(* PLC project Pump station (ladder), Digital twin lab Pump station 1 *)
(* stored: creationDateTime 2026-10-06T00:00:00, modificationDateTime 2026-10-06T00:00:00 *)

(* Lead/lag pump station control in ladder logic. Same behavior, variables and addresses as pump_station.st. *)
PROGRAM PumpStation
  VAR
    P1_RUNNING AT %IX100.0 : BOOL;  (* P1 running feedback (simulator DI 0) *)
    P2_RUNNING AT %IX100.1 : BOOL;  (* P2 running feedback (simulator DI 1) *)
    P1_FAULT AT %IX100.2 : BOOL;  (* P1 fault / trip (simulator DI 2) *)
    P2_FAULT AT %IX100.3 : BOOL;  (* P2 fault / trip (simulator DI 3) *)
    PT101_DISCH AT %IW100 : UINT;  (* Discharge pressure PT-101, psi x10 *)
    PT100_SUCT AT %IW101 : UINT;  (* Suction pressure PT-100, psi x10 *)
    DEMAND AT %IW102 : UINT;  (* Pipeline demand, % x10 *)
    SIM_HEARTBEAT AT %IW103 : UINT;  (* Simulator heartbeat, +1 every simulator step *)
    P1_RUN_CMD AT %QX100.0 : BOOL;  (* P1 run command (simulator coil 0) *)
    P2_RUN_CMD AT %QX100.1 : BOOL;  (* P2 run command (simulator coil 1) *)
    HMI_DISCH_PRESS AT %QW0 : UINT;  (* HR 0: discharge pressure, psi x10 *)
    HMI_SUCT_PRESS AT %QW1 : UINT;  (* HR 1: suction pressure, psi x10 *)
    HMI_DEMAND AT %QW2 : UINT;  (* HR 2: demand, % x10 *)
    HMI_STATUS AT %QW3 : UINT;  (* HR 3: status bits (design 5.2) *)
    HMI_ALARMS AT %QW4 : UINT;  (* HR 4: alarm bits (design 5.2) *)
    HMI_LEAD_PUMP AT %QW5 : UINT;  (* HR 5: active lead pump, 1 or 2 *)
    HMI_MODE_ACTIVE AT %QW6 : UINT;  (* HR 6: active mode, 0 Off 1 Auto 2 Manual *)
    PLC_HEARTBEAT AT %QW7 : UINT;  (* HR 7: +1 every PLC scan *)
    SP_PRESSURE AT %MW0 : UINT;  (* HR 1024: lag start pressure, psi x10 *)
    SP_LAG_STOP AT %MW1 : UINT;  (* HR 1025: lag stop pressure, psi x10 *)
    SP_LOW_ALARM AT %MW2 : UINT;  (* HR 1026: low pressure alarm, psi x10 *)
    SP_HIGH_ALARM AT %MW3 : UINT;  (* HR 1027: high pressure alarm, psi x10 *)
    LAG_START_DELAY AT %MW4 : UINT;  (* HR 1028: lag start delay, s *)
    LAG_STOP_DELAY AT %MW5 : UINT;  (* HR 1029: lag stop delay, s *)
    CMD_MODE AT %MW6 : UINT;  (* HR 1030: mode command, 0 Off 1 Auto 2 Manual *)
    CMD_LEAD_SELECT AT %MW7 : UINT;  (* HR 1031: lead pump select, 1 = P1, 2 = P2 *)
    CMD_MANUAL_P1 AT %MW8 : UINT;  (* HR 1032: Manual mode P1, 1 run 0 stop *)
    CMD_MANUAL_P2 AT %MW9 : UINT;  (* HR 1033: Manual mode P2, 1 run 0 stop *)
    CMD_ALARM_RESET AT %MW10 : UINT;  (* HR 1034: alarm reset, HMI writes 1, PLC clears it *)
  END_VAR
  VAR
    LoadDefaults : BOOL;  (* SP_PRESSURE is 0: settings were never written, load defaults *)
    MinLagStop : UINT;  (* SP_PRESSURE + 10 psi, the lowest allowed lag stop pressure *)
    ModeAuto : BOOL;  (* CMD_MODE = 1 *)
    ModeManual : BOOL;  (* CMD_MODE = 2 *)
    SelP2 : BOOL;  (* CMD_LEAD_SELECT = 2 (operator wants P2 as lead) *)
    ManP1 : BOOL;  (* CMD_MANUAL_P1 = 1 *)
    ManP2 : BOOL;  (* CMD_MANUAL_P2 = 1 *)
    ResetReq : BOOL;  (* Operator pressed Reset (CMD_ALARM_RESET <> 0) *)
    PressBelowSP : BOOL;  (* Discharge pressure below the lag start pressure *)
    PressAboveLagStop : BOOL;  (* Discharge pressure above the lag stop pressure *)
    PressBelowLowAlm : BOOL;  (* Discharge pressure below the low alarm limit *)
    PressAboveHighAlm : BOOL;  (* Discharge pressure above the high alarm limit *)
    P1StartTmr : TON;  (* P1 commanded but not running *)
    P2StartTmr : TON;  (* P2 commanded but not running *)
    P1StartFail : BOOL;  (* P1 failed to start within 5 s *)
    P2StartFail : BOOL;  (* P2 failed to start within 5 s *)
    P1Failed : BOOL;  (* P1 locked out (fault or failed to start) until Reset *)
    P2Failed : BOOL;  (* P2 locked out (fault or failed to start) until Reset *)
    EnterAuto : BOOL;  (* First scan in Auto *)
    LeadIsP2 : BOOL;  (* Active lead pump: FALSE = P1, TRUE = P2 (ActiveLead in the ST program) *)
    LagPumpCmd : BOOL;  (* The pump that is now lag is commanded to run *)
    FailToP2 : BOOL;  (* Lead P1 has failed and P2 is healthy: make P2 lead *)
    FailToP1 : BOOL;  (* Lead P2 has failed and P1 is healthy: make P1 lead *)
    LeadChange : BOOL;  (* Apply the operator's new lead selection this scan *)
    LagRun : BOOL;  (* Auto logic wants the lag pump running *)
    Handover : BOOL;  (* Lead change in progress: old lead keeps running until the new one runs *)
    LeadAvail : BOOL;  (* Lead pump is not locked out *)
    LagAvail : BOOL;  (* Lag pump is not locked out *)
    LeadRunning : BOOL;  (* Lead pump reports running *)
    LagStartPT : TIME;  (* Lag start delay as TIME *)
    LagStopPT : TIME;  (* Lag stop delay as TIME *)
    LagStartTmr : TON;  (* Pressure low long enough to start the lag pump *)
    LagStopTmr : TON;  (* Pressure high long enough to stop the lag pump *)
    LagStartDone : BOOL;  (* LagStartTmr.Q *)
    LagStopDone : BOOL;  (* LagStopTmr.Q *)
    LowArmTmr : TON;  (* Start-up bypass for the low pressure alarm *)
    LowPressTmr : TON;  (* Low pressure alarm delay *)
    HighPressTmr : TON;  (* High pressure alarm delay *)
    CommLossTmr : TON;  (* Simulator heartbeat frozen *)
    LowArmed : BOOL;  (* Low pressure alarm armed (15 s out of Off) *)
    LowPressOn : BOOL;  (* Pressure low for 5 s *)
    HighPressOn : BOOL;  (* Pressure high for 5 s *)
    SimHbFrozen : BOOL;  (* Simulator heartbeat unchanged since the last scan *)
    LastSimHb : UINT;  (* Simulator heartbeat seen last scan *)
    CommLost : BOOL;  (* Simulator heartbeat frozen for 3 s *)
    CommOk : BOOL;  (* Simulator link healthy *)
    AlmLow : BOOL;  (* Low discharge pressure alarm (latched) *)
    AlmHigh : BOOL;  (* High discharge pressure alarm (latched) *)
    AlmComm : BOOL;  (* Simulator comm loss alarm (latched) *)
    AlmUnack : BOOL;  (* A new alarm has not been acknowledged *)
    AnyAlarm : BOOL;  (* Any alarm or pump lockout active *)
    LagRunning : BOOL;  (* Lag pump reports running *)
    StatusWord : UINT;  (* HMI_STATUS being built *)
    AlarmWord : UINT;  (* HMI_ALARMS being built *)
    HbWrap : BOOL;  (* PLC_HEARTBEAT is at 65535 and wraps to 0 *)
  END_VAR
  VAR  (* added by the conversion: wires and edge detectors of the diagram *)
    R_TRIG1 : R_TRIG;
    R_TRIG2 : R_TRIG;
  END_VAR

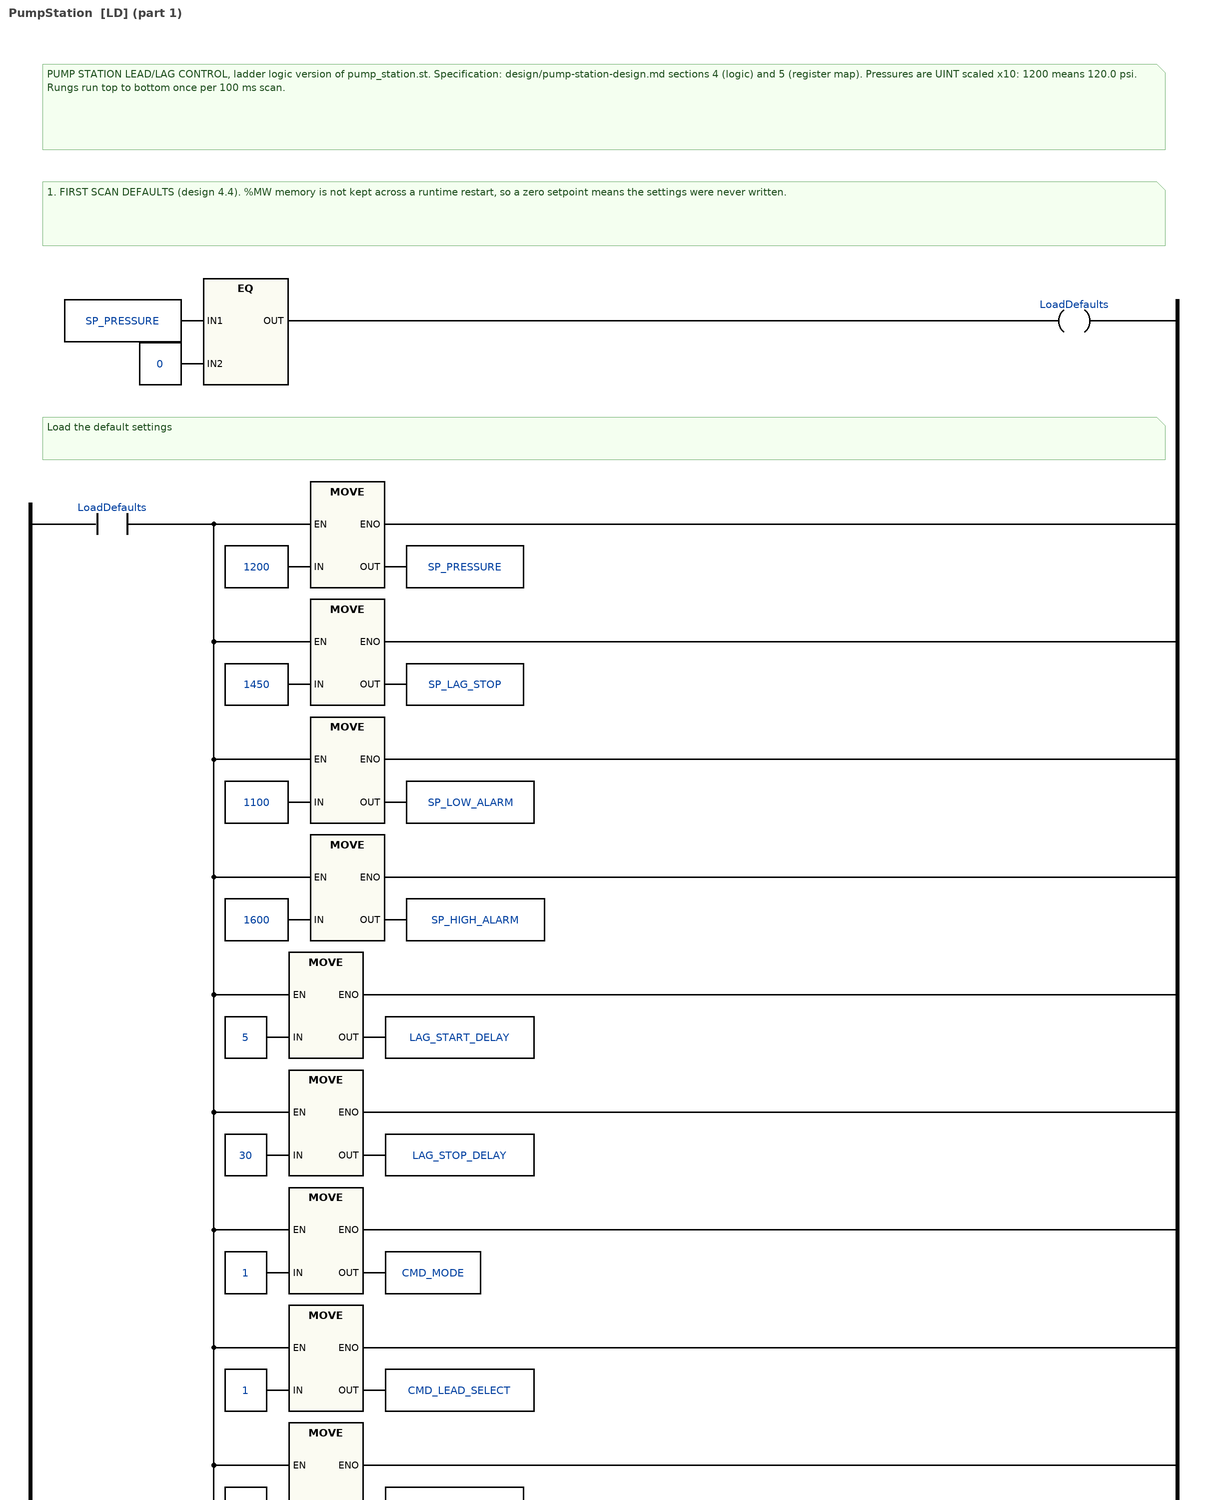
(* LD diagram, written out as Structured Text *)
(* PUMP STATION LEAD/LAG CONTROL, ladder logic version of pump_station.st. Specification: design/pump-station-design.md sections 4 (logic) and 5 (register map). Pressures are UINT scaled x10: 1200 means 120.0 psi. Rungs run top to bottom once per 100 ms scan. *)
(* 1. FIRST SCAN DEFAULTS (design 4.4). %MW memory is not kept across a runtime restart, so a zero setpoint means the settings were never written. *)
LoadDefaults := SP_PRESSURE = 0;
(* Load the default settings *)
IF LoadDefaults THEN SP_PRESSURE := 1200; END_IF;
IF LoadDefaults THEN SP_LAG_STOP := 1450; END_IF;
IF LoadDefaults THEN SP_LOW_ALARM := 1100; END_IF;
IF LoadDefaults THEN SP_HIGH_ALARM := 1600; END_IF;
IF LoadDefaults THEN LAG_START_DELAY := 5; END_IF;
IF LoadDefaults THEN LAG_STOP_DELAY := 30; END_IF;
IF LoadDefaults THEN CMD_MODE := 1; END_IF;
IF LoadDefaults THEN CMD_LEAD_SELECT := 1; END_IF;
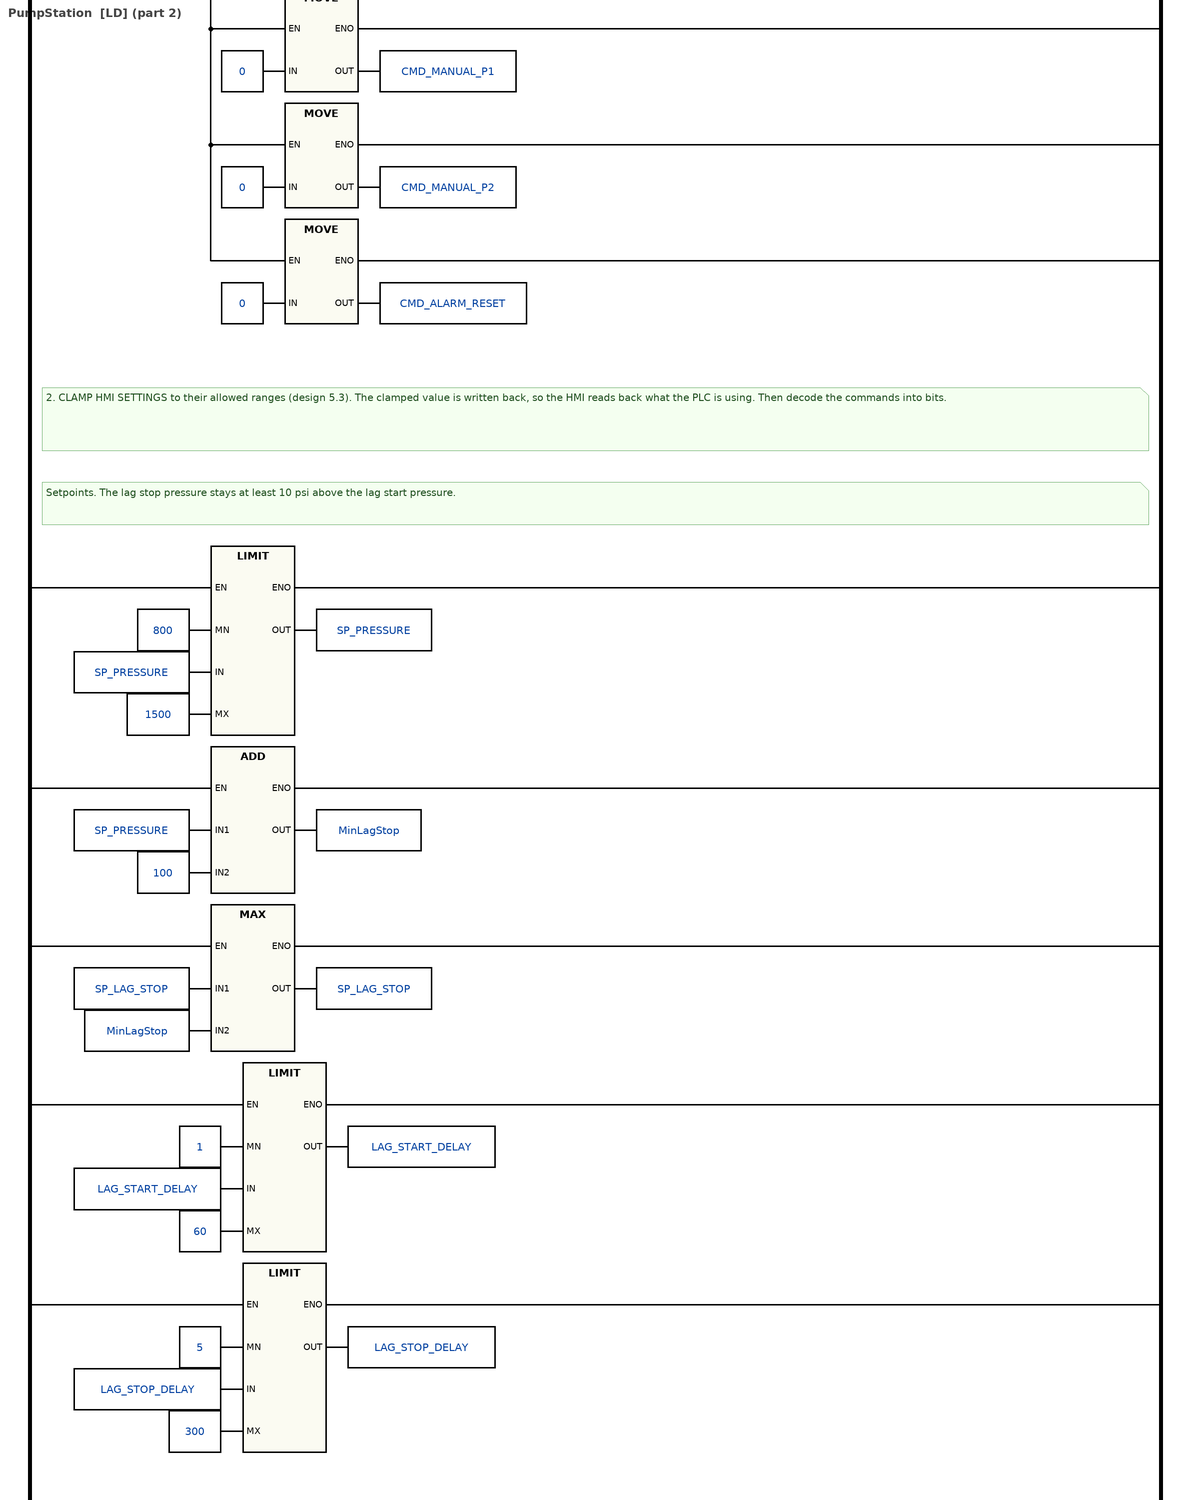
IF LoadDefaults THEN CMD_MANUAL_P1 := 0; END_IF;
IF LoadDefaults THEN CMD_MANUAL_P2 := 0; END_IF;
IF LoadDefaults THEN CMD_ALARM_RESET := 0; END_IF;
(* 2. CLAMP HMI SETTINGS to their allowed ranges (design 5.3). The clamped value is written back, so the HMI reads back what the PLC is using. Then decode the commands into bits. *)
(* Setpoints. The lag stop pressure stays at least 10 psi above the lag start pressure. *)
SP_PRESSURE := LIMIT(800, SP_PRESSURE, 1500);
MinLagStop := SP_PRESSURE + 100;
SP_LAG_STOP := MAX(SP_LAG_STOP, MinLagStop);
LAG_START_DELAY := LIMIT(1, LAG_START_DELAY, 60);
LAG_STOP_DELAY := LIMIT(5, LAG_STOP_DELAY, 300);
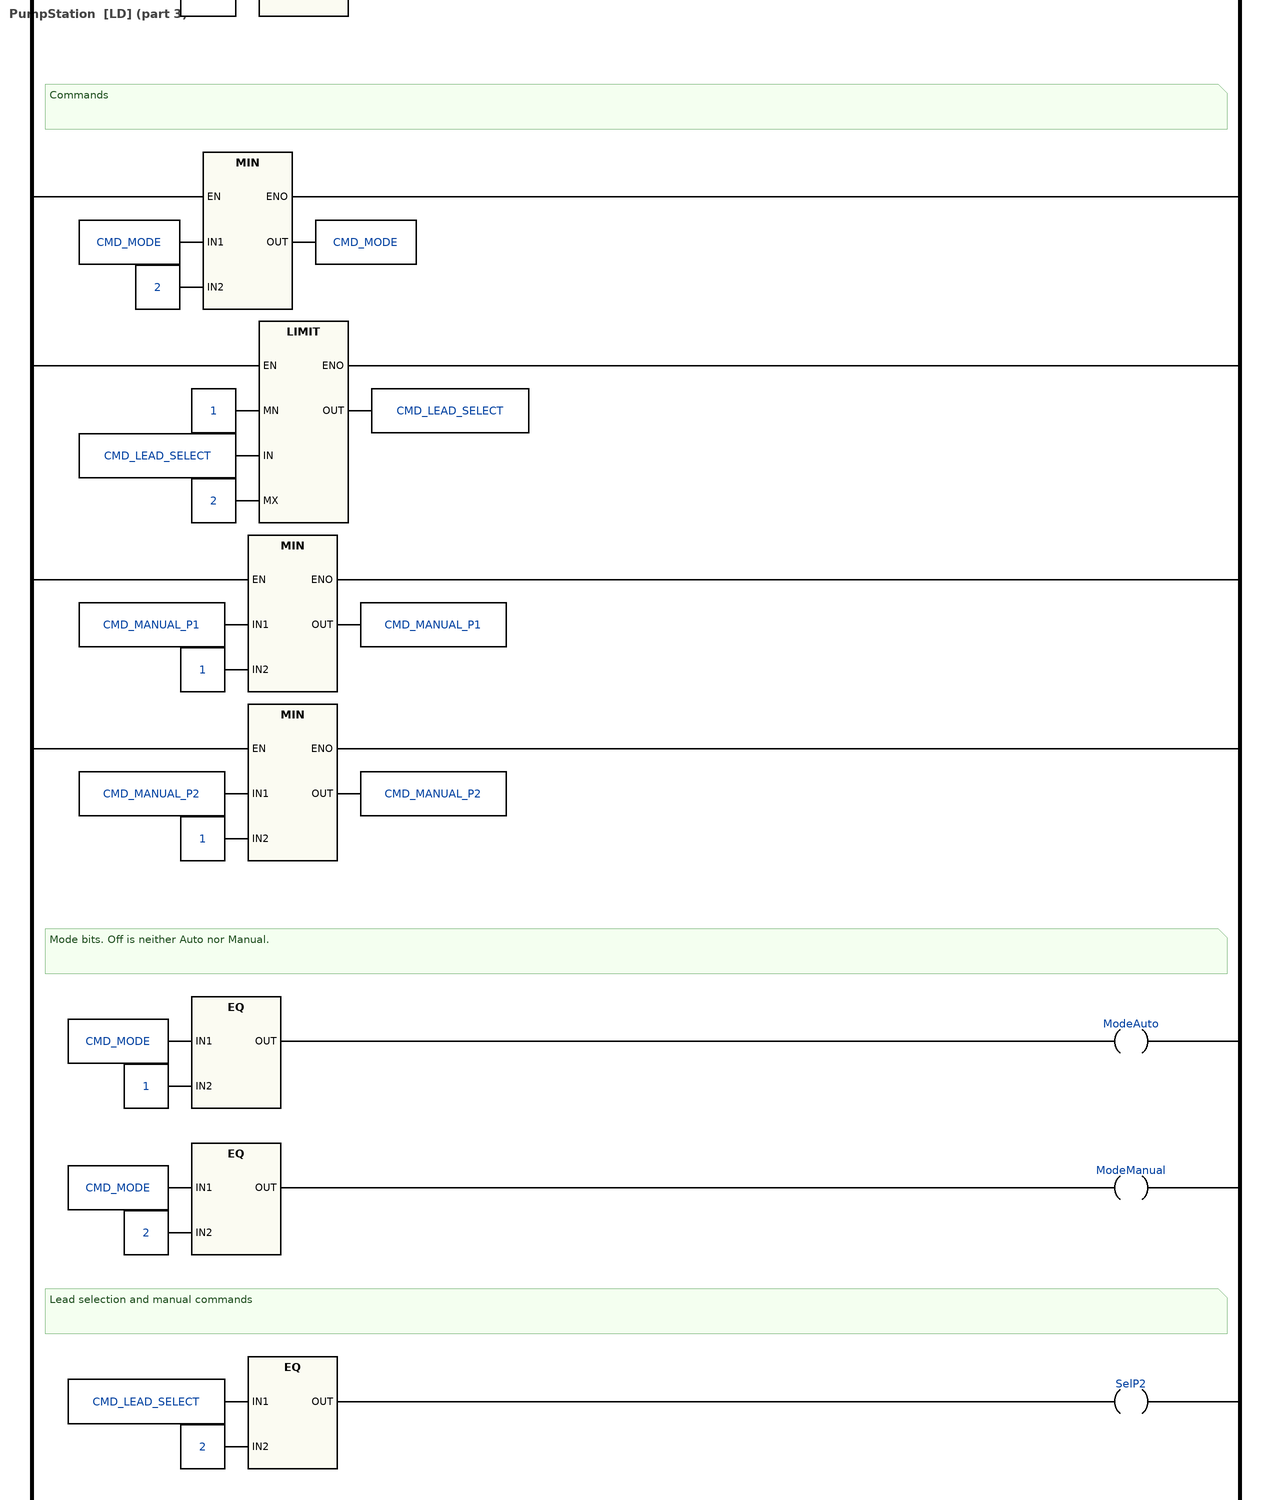
(* Commands *)
CMD_MODE := MIN(CMD_MODE, 2);
CMD_LEAD_SELECT := LIMIT(1, CMD_LEAD_SELECT, 2);
CMD_MANUAL_P1 := MIN(CMD_MANUAL_P1, 1);
CMD_MANUAL_P2 := MIN(CMD_MANUAL_P2, 1);
(* Mode bits. Off is neither Auto nor Manual. *)
ModeAuto := CMD_MODE = 1;
ModeManual := CMD_MODE = 2;
(* Lead selection and manual commands *)
SelP2 := CMD_LEAD_SELECT = 2;
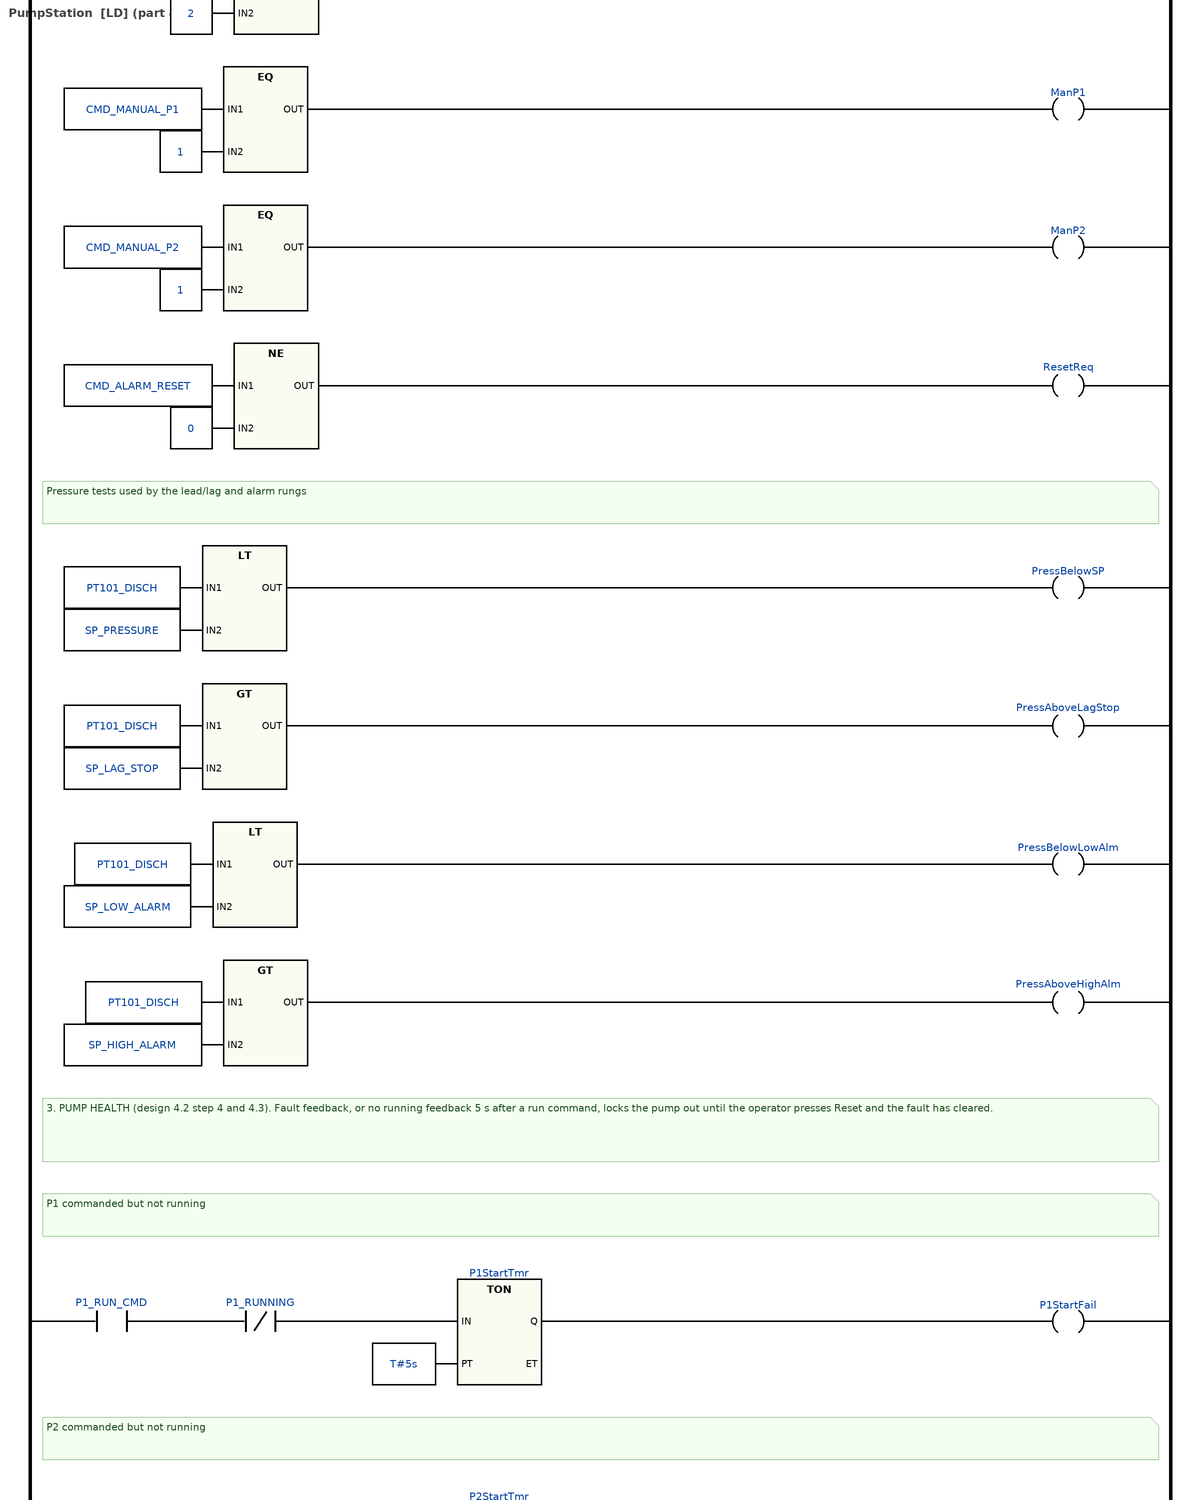
ManP1 := CMD_MANUAL_P1 = 1;
ManP2 := CMD_MANUAL_P2 = 1;
ResetReq := CMD_ALARM_RESET <> 0;
(* Pressure tests used by the lead/lag and alarm rungs *)
PressBelowSP := PT101_DISCH < SP_PRESSURE;
PressAboveLagStop := PT101_DISCH > SP_LAG_STOP;
PressBelowLowAlm := PT101_DISCH < SP_LOW_ALARM;
PressAboveHighAlm := PT101_DISCH > SP_HIGH_ALARM;
(* 3. PUMP HEALTH (design 4.2 step 4 and 4.3). Fault feedback, or no running feedback 5 s after a run command, locks the pump out until the operator presses Reset and the fault has cleared. *)
(* P1 commanded but not running *)
P1StartTmr(IN := P1_RUN_CMD AND NOT P1_RUNNING, PT := T#5s);
P1StartFail := P1StartTmr.Q;
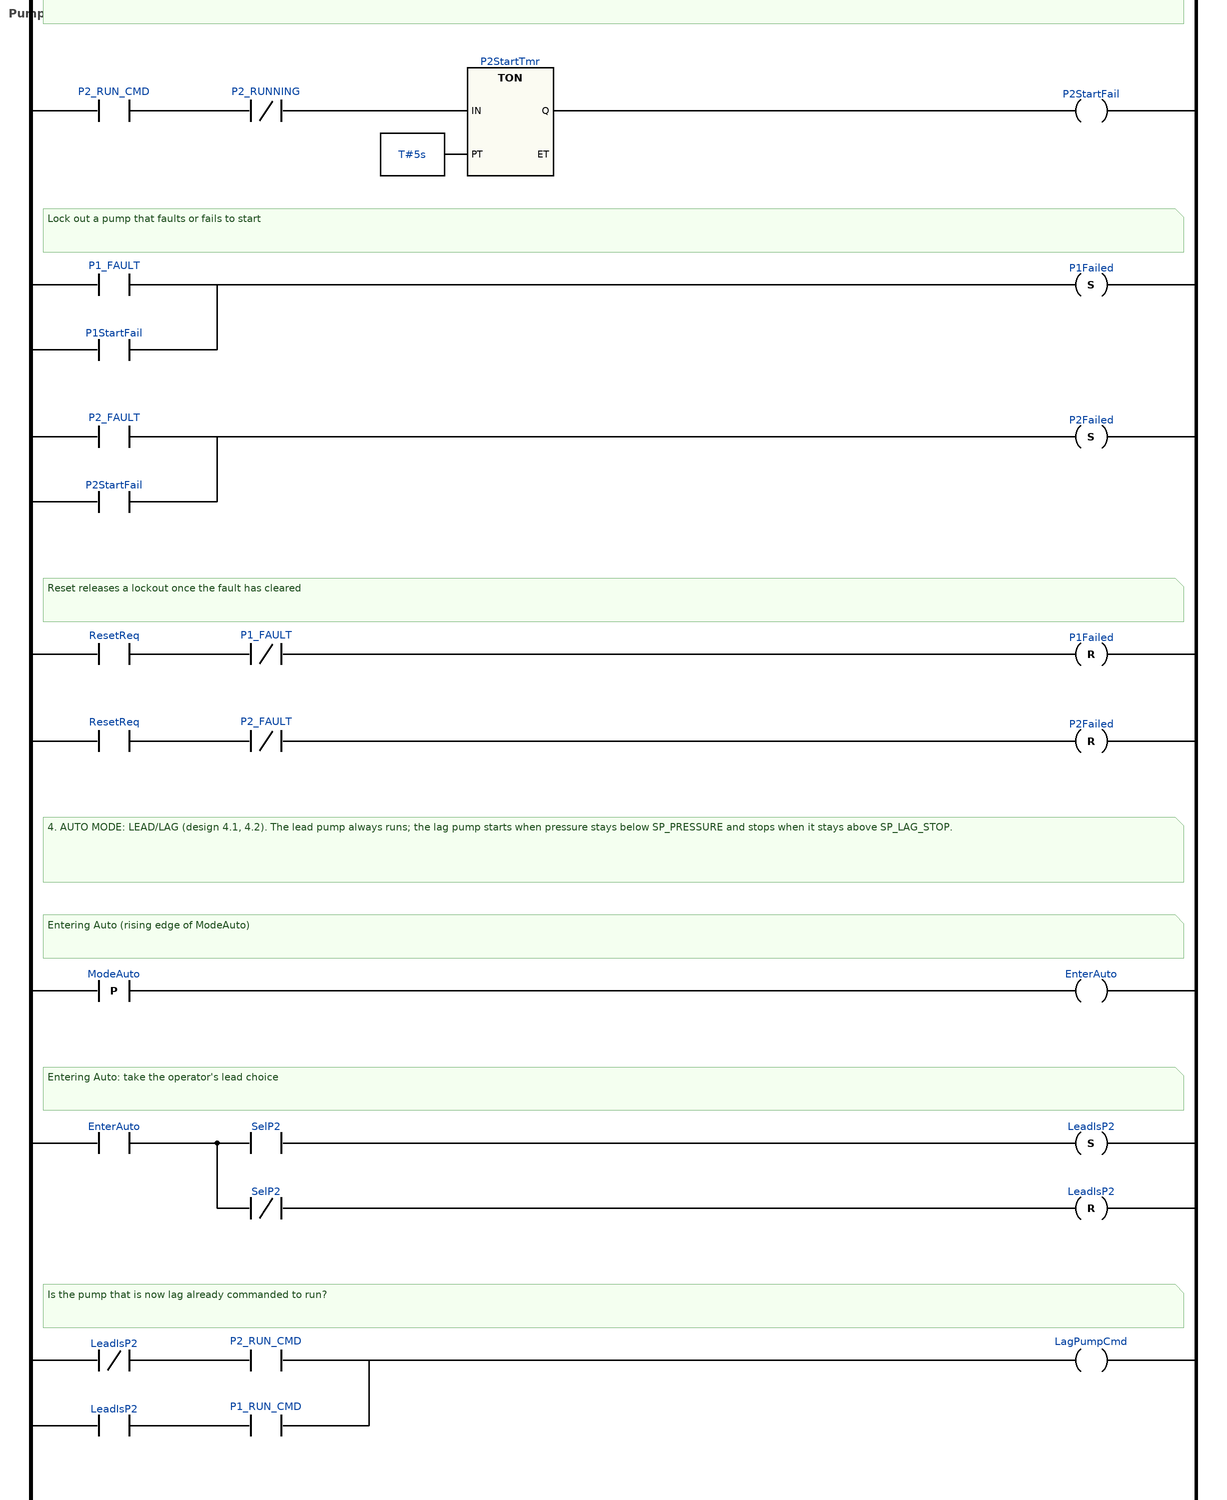
(* P2 commanded but not running *)
P2StartTmr(IN := P2_RUN_CMD AND NOT P2_RUNNING, PT := T#5s);
P2StartFail := P2StartTmr.Q;
(* Lock out a pump that faults or fails to start *)
IF P1_FAULT OR P1StartFail THEN P1Failed := TRUE; END_IF;
IF P2_FAULT OR P2StartFail THEN P2Failed := TRUE; END_IF;
(* Reset releases a lockout once the fault has cleared *)
IF ResetReq AND NOT P1_FAULT THEN P1Failed := FALSE; END_IF;
IF ResetReq AND NOT P2_FAULT THEN P2Failed := FALSE; END_IF;
(* 4. AUTO MODE: LEAD/LAG (design 4.1, 4.2). The lead pump always runs; the lag pump starts when pressure stays below SP_PRESSURE and stops when it stays above SP_LAG_STOP. *)
(* Entering Auto (rising edge of ModeAuto) *)
R_TRIG1(CLK := ModeAuto);
EnterAuto := R_TRIG1.Q;
(* Entering Auto: take the operator's lead choice *)
IF EnterAuto AND SelP2 THEN LeadIsP2 := TRUE; END_IF;
IF EnterAuto AND NOT SelP2 THEN LeadIsP2 := FALSE; END_IF;
(* Is the pump that is now lag already commanded to run? *)
LagPumpCmd := NOT LeadIsP2 AND P2_RUN_CMD OR LeadIsP2 AND P1_RUN_CMD;
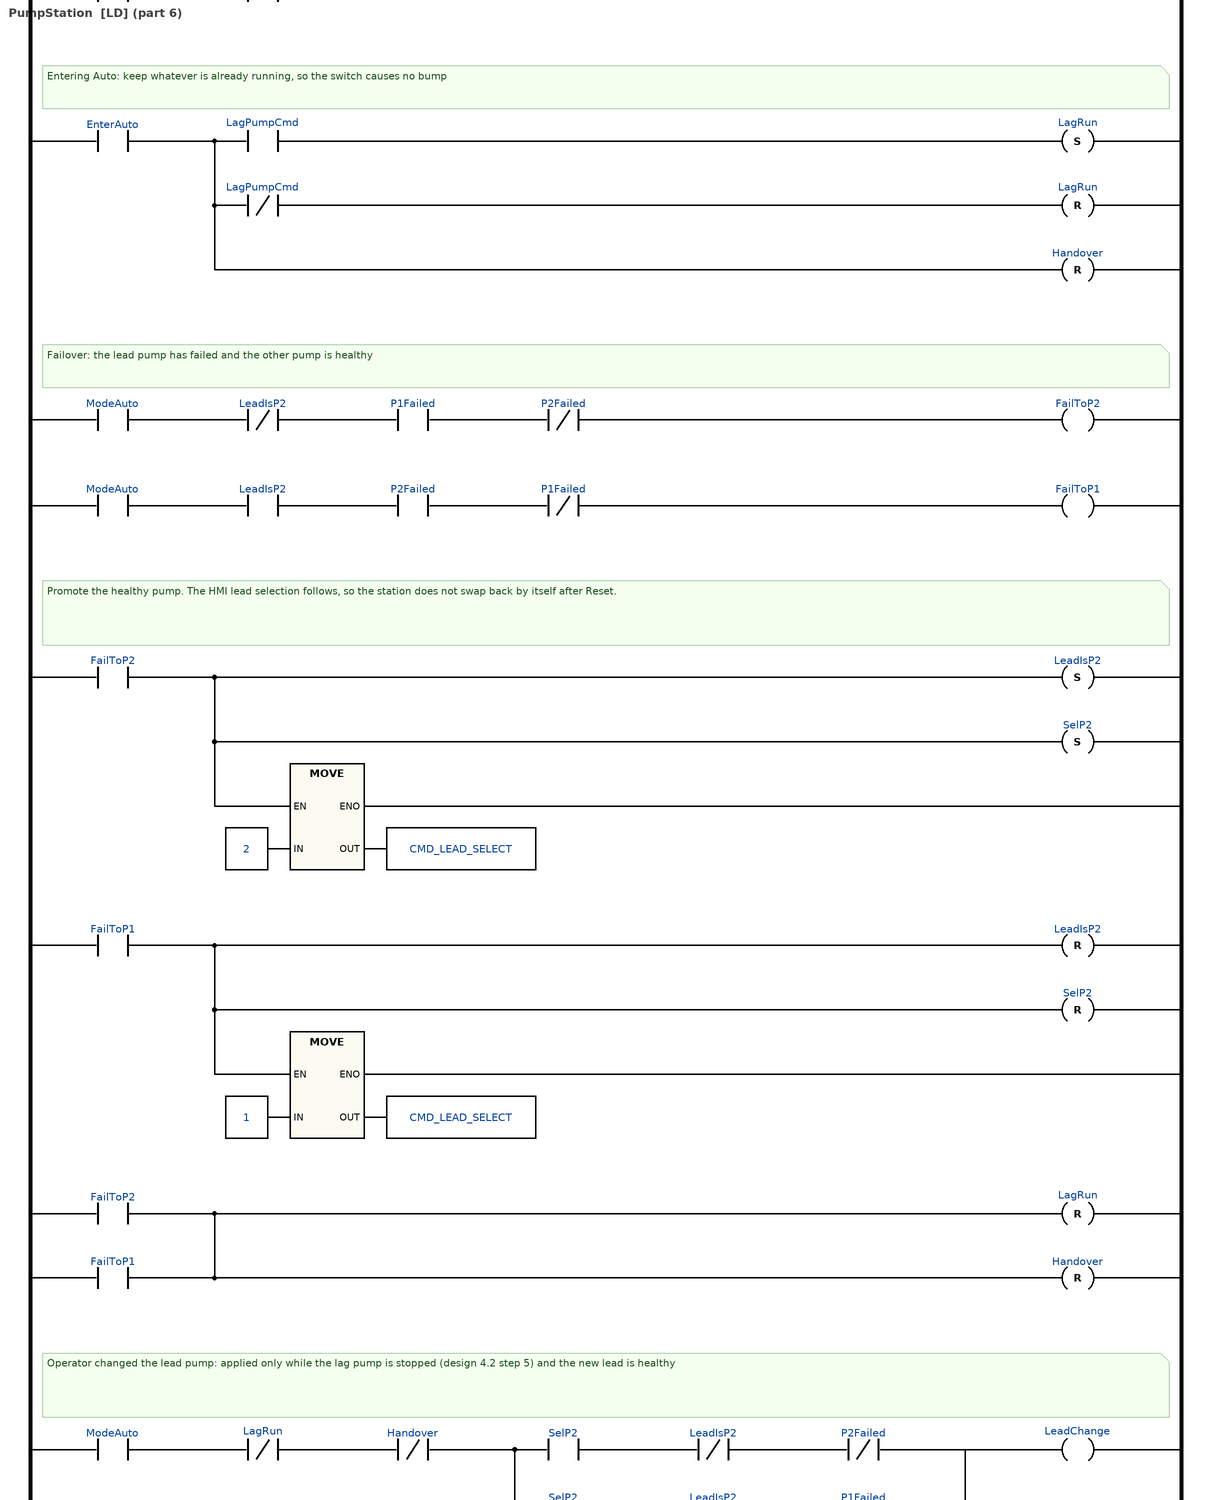
(* Entering Auto: keep whatever is already running, so the switch causes no bump *)
IF EnterAuto AND LagPumpCmd THEN LagRun := TRUE; END_IF;
IF EnterAuto AND NOT LagPumpCmd THEN LagRun := FALSE; END_IF;
IF EnterAuto THEN Handover := FALSE; END_IF;
(* Failover: the lead pump has failed and the other pump is healthy *)
FailToP2 := ModeAuto AND NOT LeadIsP2 AND P1Failed AND NOT P2Failed;
FailToP1 := ModeAuto AND LeadIsP2 AND P2Failed AND NOT P1Failed;
(* Promote the healthy pump. The HMI lead selection follows, so the station does not swap back by itself after Reset. *)
IF FailToP2 THEN LeadIsP2 := TRUE; END_IF;
IF FailToP2 THEN SelP2 := TRUE; END_IF;
IF FailToP2 THEN CMD_LEAD_SELECT := 2; END_IF;
IF FailToP1 THEN LeadIsP2 := FALSE; END_IF;
IF FailToP1 THEN SelP2 := FALSE; END_IF;
IF FailToP1 THEN CMD_LEAD_SELECT := 1; END_IF;
IF FailToP2 OR FailToP1 THEN LagRun := FALSE; END_IF;
IF FailToP2 OR FailToP1 THEN Handover := FALSE; END_IF;
(* Operator changed the lead pump: applied only while the lag pump is stopped (design 4.2 step 5) and the new lead is healthy *)
LeadChange := ModeAuto AND NOT LagRun AND NOT Handover AND (SelP2 AND NOT LeadIsP2 AND NOT P2Failed OR NOT SelP2 AND LeadIsP2 AND NOT P1Failed);
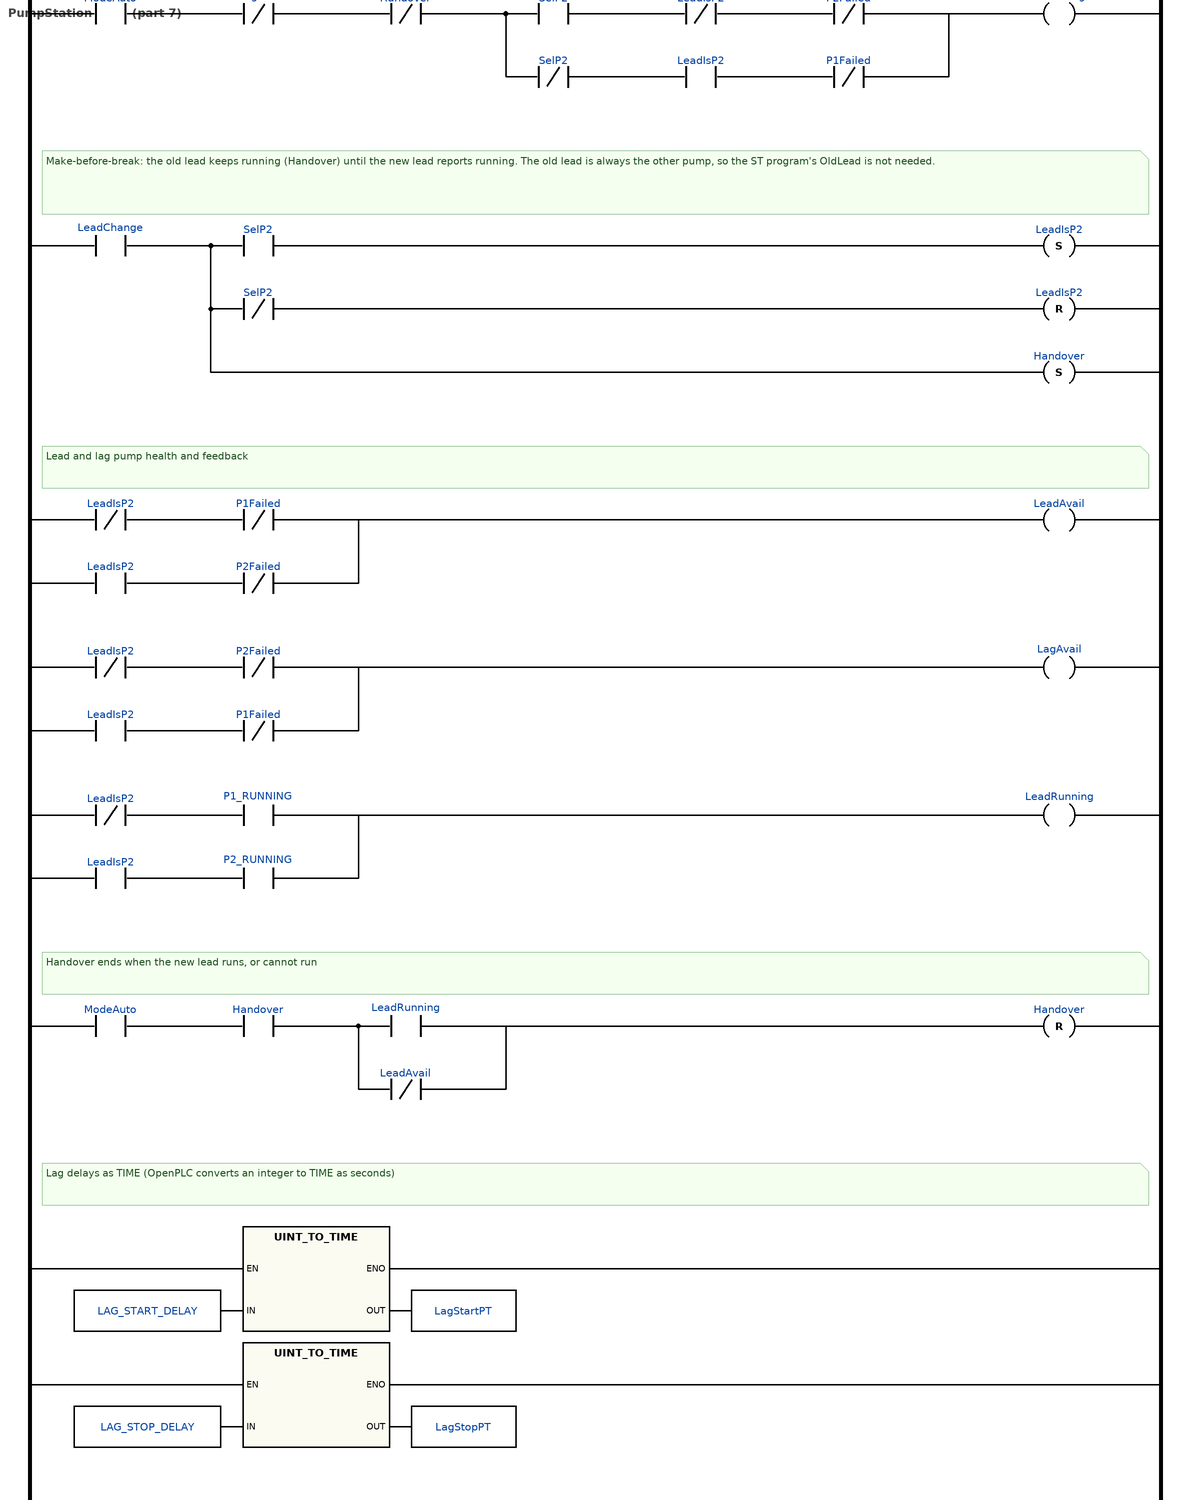
(* Make-before-break: the old lead keeps running (Handover) until the new lead reports running. The old lead is always the other pump, so the ST program's OldLead is not needed. *)
IF LeadChange AND SelP2 THEN LeadIsP2 := TRUE; END_IF;
IF LeadChange AND NOT SelP2 THEN LeadIsP2 := FALSE; END_IF;
IF LeadChange THEN Handover := TRUE; END_IF;
(* Lead and lag pump health and feedback *)
LeadAvail := NOT LeadIsP2 AND NOT P1Failed OR LeadIsP2 AND NOT P2Failed;
LagAvail := NOT LeadIsP2 AND NOT P2Failed OR LeadIsP2 AND NOT P1Failed;
LeadRunning := NOT LeadIsP2 AND P1_RUNNING OR LeadIsP2 AND P2_RUNNING;
(* Handover ends when the new lead runs, or cannot run *)
IF ModeAuto AND Handover AND (LeadRunning OR NOT LeadAvail) THEN Handover := FALSE; END_IF;
(* Lag delays as TIME (OpenPLC converts an integer to TIME as seconds) *)
LagStartPT := UINT_TO_TIME(LAG_START_DELAY);
LagStopPT := UINT_TO_TIME(LAG_STOP_DELAY);
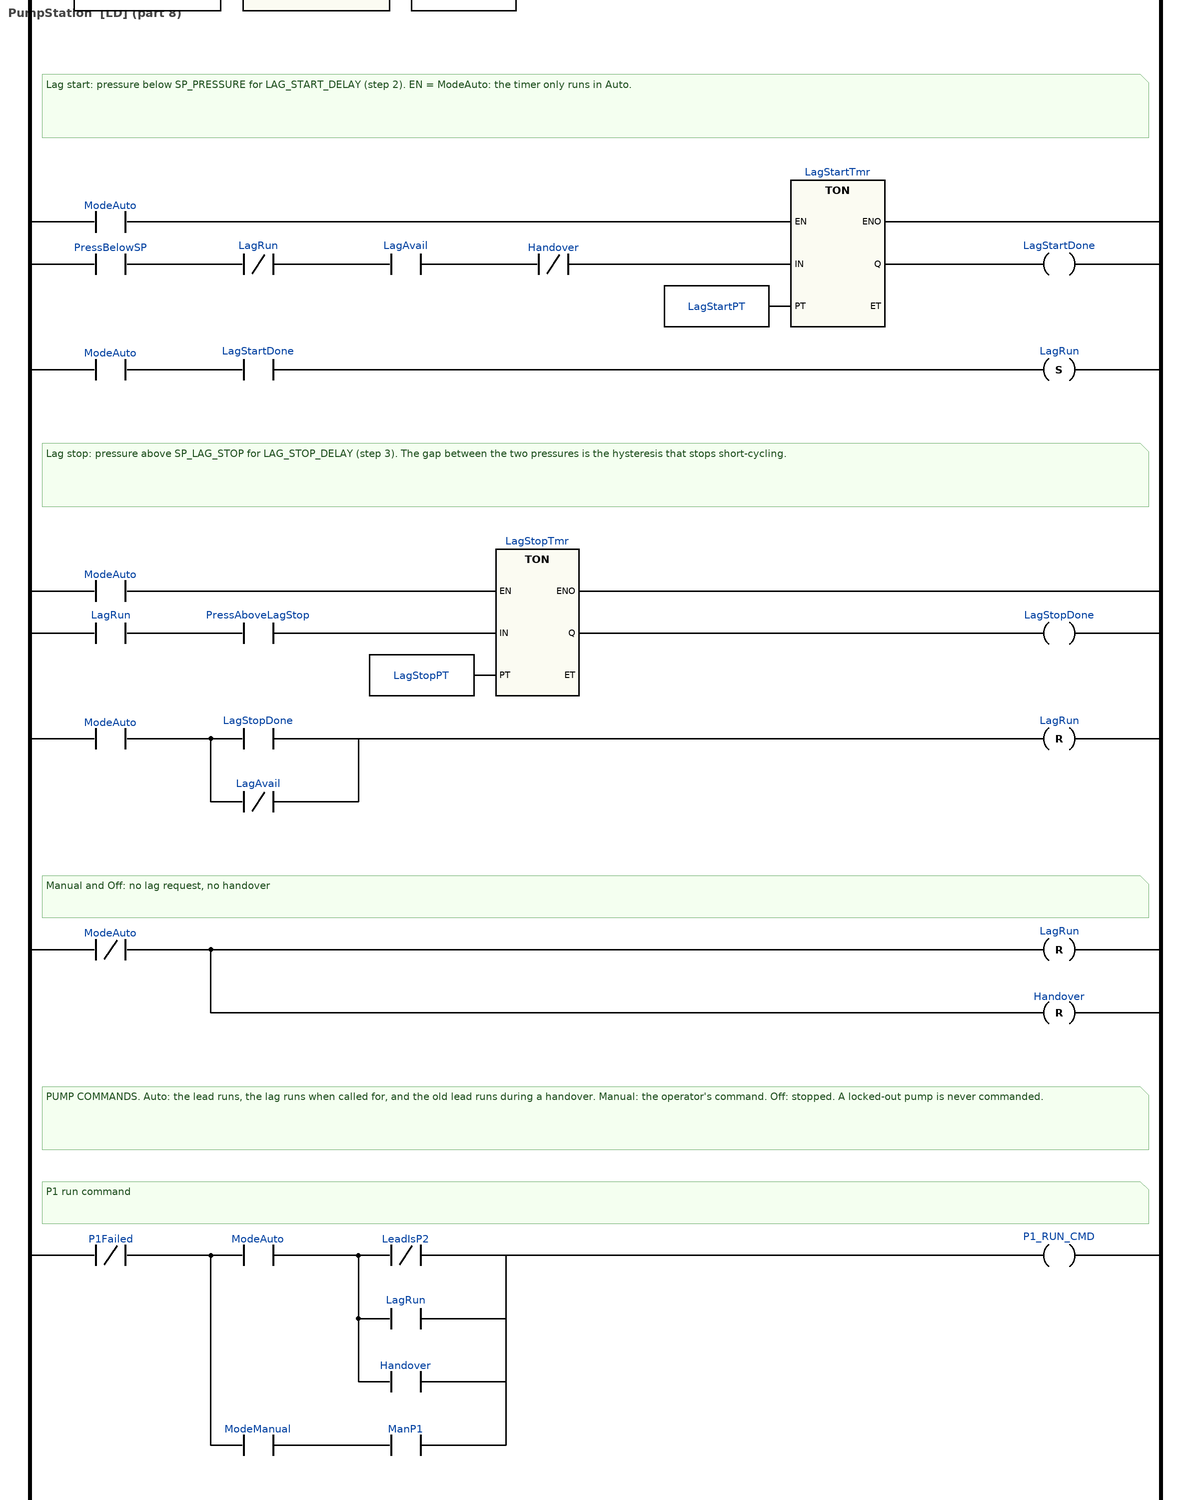
(* Lag start: pressure below SP_PRESSURE for LAG_START_DELAY (step 2). EN = ModeAuto: the timer only runs in Auto. *)
LagStartTmr(EN := ModeAuto, IN := PressBelowSP AND NOT LagRun AND LagAvail AND NOT Handover, PT := LagStartPT);
LagStartDone := LagStartTmr.Q;
IF ModeAuto AND LagStartDone THEN LagRun := TRUE; END_IF;
(* Lag stop: pressure above SP_LAG_STOP for LAG_STOP_DELAY (step 3). The gap between the two pressures is the hysteresis that stops short-cycling. *)
LagStopTmr(EN := ModeAuto, IN := LagRun AND PressAboveLagStop, PT := LagStopPT);
LagStopDone := LagStopTmr.Q;
IF ModeAuto AND (LagStopDone OR NOT LagAvail) THEN LagRun := FALSE; END_IF;
(* Manual and Off: no lag request, no handover *)
IF NOT ModeAuto THEN LagRun := FALSE; END_IF;
IF NOT ModeAuto THEN Handover := FALSE; END_IF;
(* PUMP COMMANDS. Auto: the lead runs, the lag runs when called for, and the old lead runs during a handover. Manual: the operator's command. Off: stopped. A locked-out pump is never commanded. *)
(* P1 run command *)
P1_RUN_CMD := NOT P1Failed AND (ModeAuto AND NOT LeadIsP2 OR ModeAuto AND LagRun OR ModeAuto AND Handover OR ModeManual AND ManP1);
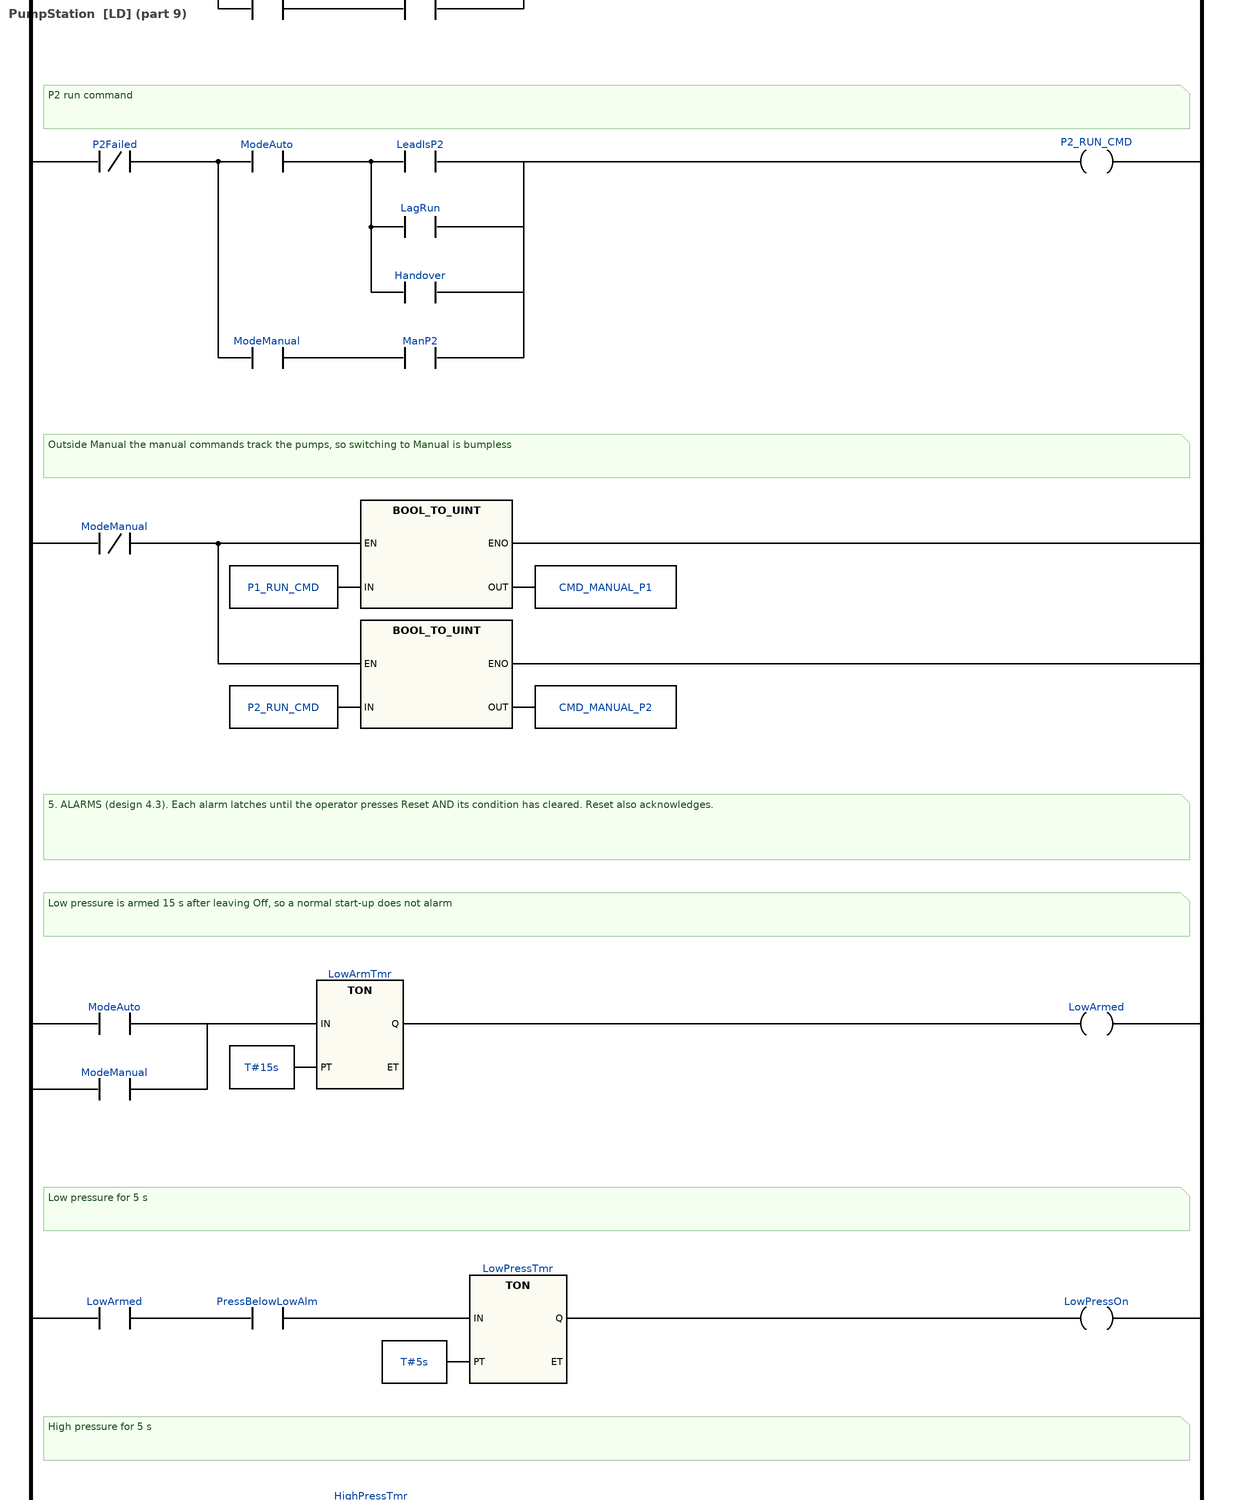
(* P2 run command *)
P2_RUN_CMD := NOT P2Failed AND (ModeAuto AND LeadIsP2 OR ModeAuto AND LagRun OR ModeAuto AND Handover OR ModeManual AND ManP2);
(* Outside Manual the manual commands track the pumps, so switching to Manual is bumpless *)
IF NOT ModeManual THEN CMD_MANUAL_P1 := BOOL_TO_UINT(P1_RUN_CMD); END_IF;
IF NOT ModeManual THEN CMD_MANUAL_P2 := BOOL_TO_UINT(P2_RUN_CMD); END_IF;
(* 5. ALARMS (design 4.3). Each alarm latches until the operator presses Reset AND its condition has cleared. Reset also acknowledges. *)
(* Low pressure is armed 15 s after leaving Off, so a normal start-up does not alarm *)
LowArmTmr(IN := ModeAuto OR ModeManual, PT := T#15s);
LowArmed := LowArmTmr.Q;
(* Low pressure for 5 s *)
LowPressTmr(IN := LowArmed AND PressBelowLowAlm, PT := T#5s);
LowPressOn := LowPressTmr.Q;
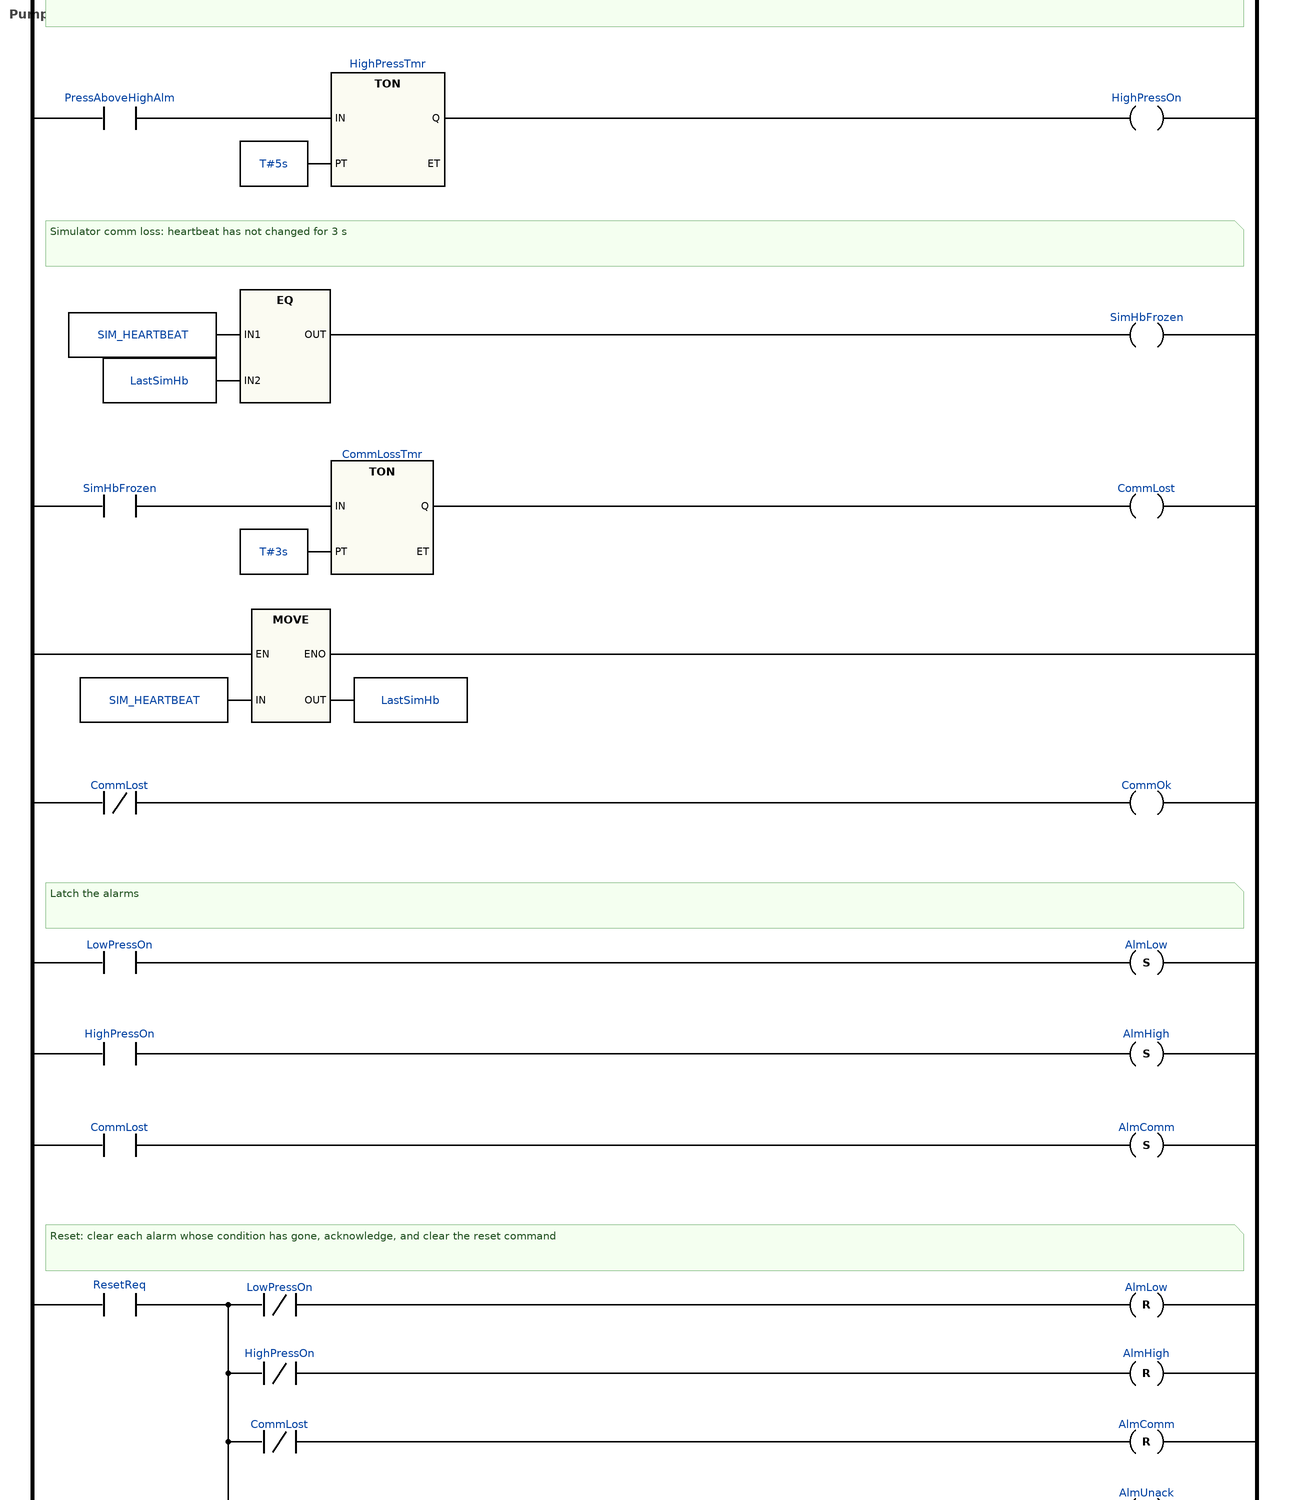
(* High pressure for 5 s *)
HighPressTmr(IN := PressAboveHighAlm, PT := T#5s);
HighPressOn := HighPressTmr.Q;
(* Simulator comm loss: heartbeat has not changed for 3 s *)
SimHbFrozen := SIM_HEARTBEAT = LastSimHb;
CommLossTmr(IN := SimHbFrozen, PT := T#3s);
CommLost := CommLossTmr.Q;
LastSimHb := SIM_HEARTBEAT;
CommOk := NOT CommLost;
(* Latch the alarms *)
IF LowPressOn THEN AlmLow := TRUE; END_IF;
IF HighPressOn THEN AlmHigh := TRUE; END_IF;
IF CommLost THEN AlmComm := TRUE; END_IF;
(* Reset: clear each alarm whose condition has gone, acknowledge, and clear the reset command *)
IF ResetReq AND NOT LowPressOn THEN AlmLow := FALSE; END_IF;
IF ResetReq AND NOT HighPressOn THEN AlmHigh := FALSE; END_IF;
IF ResetReq AND NOT CommLost THEN AlmComm := FALSE; END_IF;
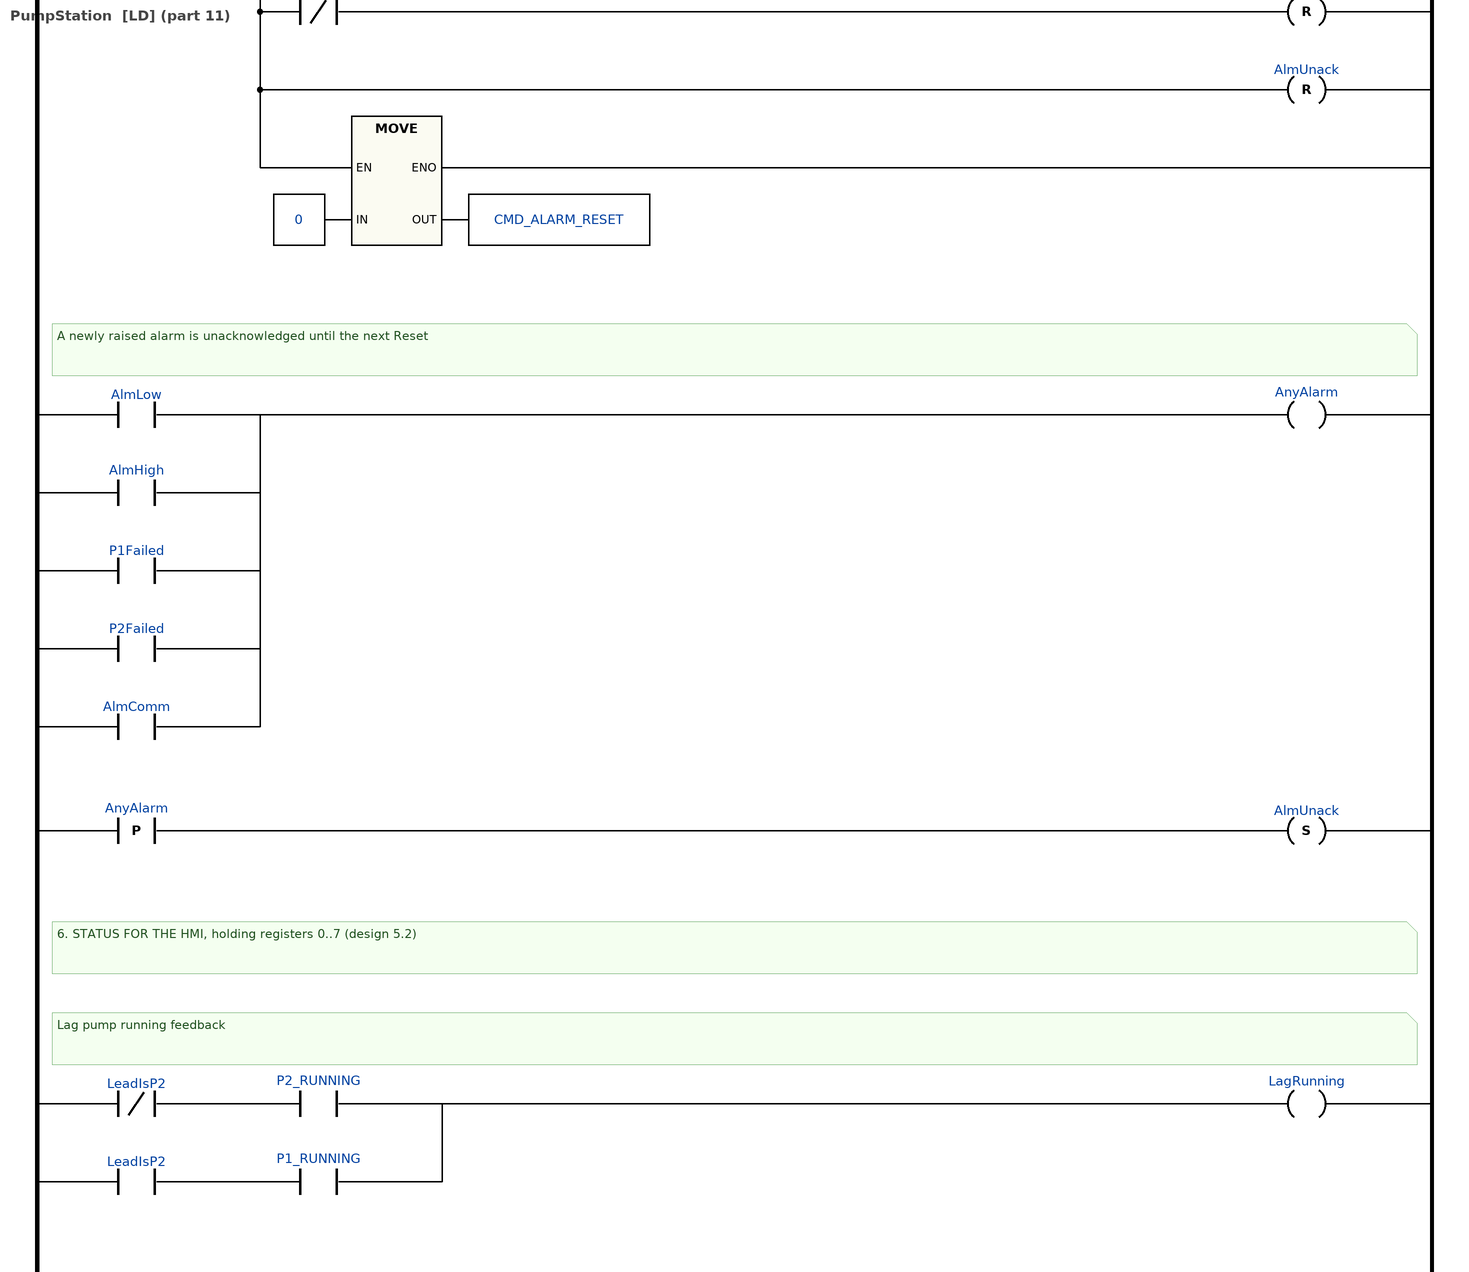
IF ResetReq THEN AlmUnack := FALSE; END_IF;
IF ResetReq THEN CMD_ALARM_RESET := 0; END_IF;
(* A newly raised alarm is unacknowledged until the next Reset *)
AnyAlarm := AlmLow OR AlmHigh OR P1Failed OR P2Failed OR AlmComm;
R_TRIG2(CLK := AnyAlarm);
IF R_TRIG2.Q THEN AlmUnack := TRUE; END_IF;
(* 6. STATUS FOR THE HMI, holding registers 0..7 (design 5.2) *)
(* Lag pump running feedback *)
LagRunning := NOT LeadIsP2 AND P2_RUNNING OR LeadIsP2 AND P1_RUNNING;
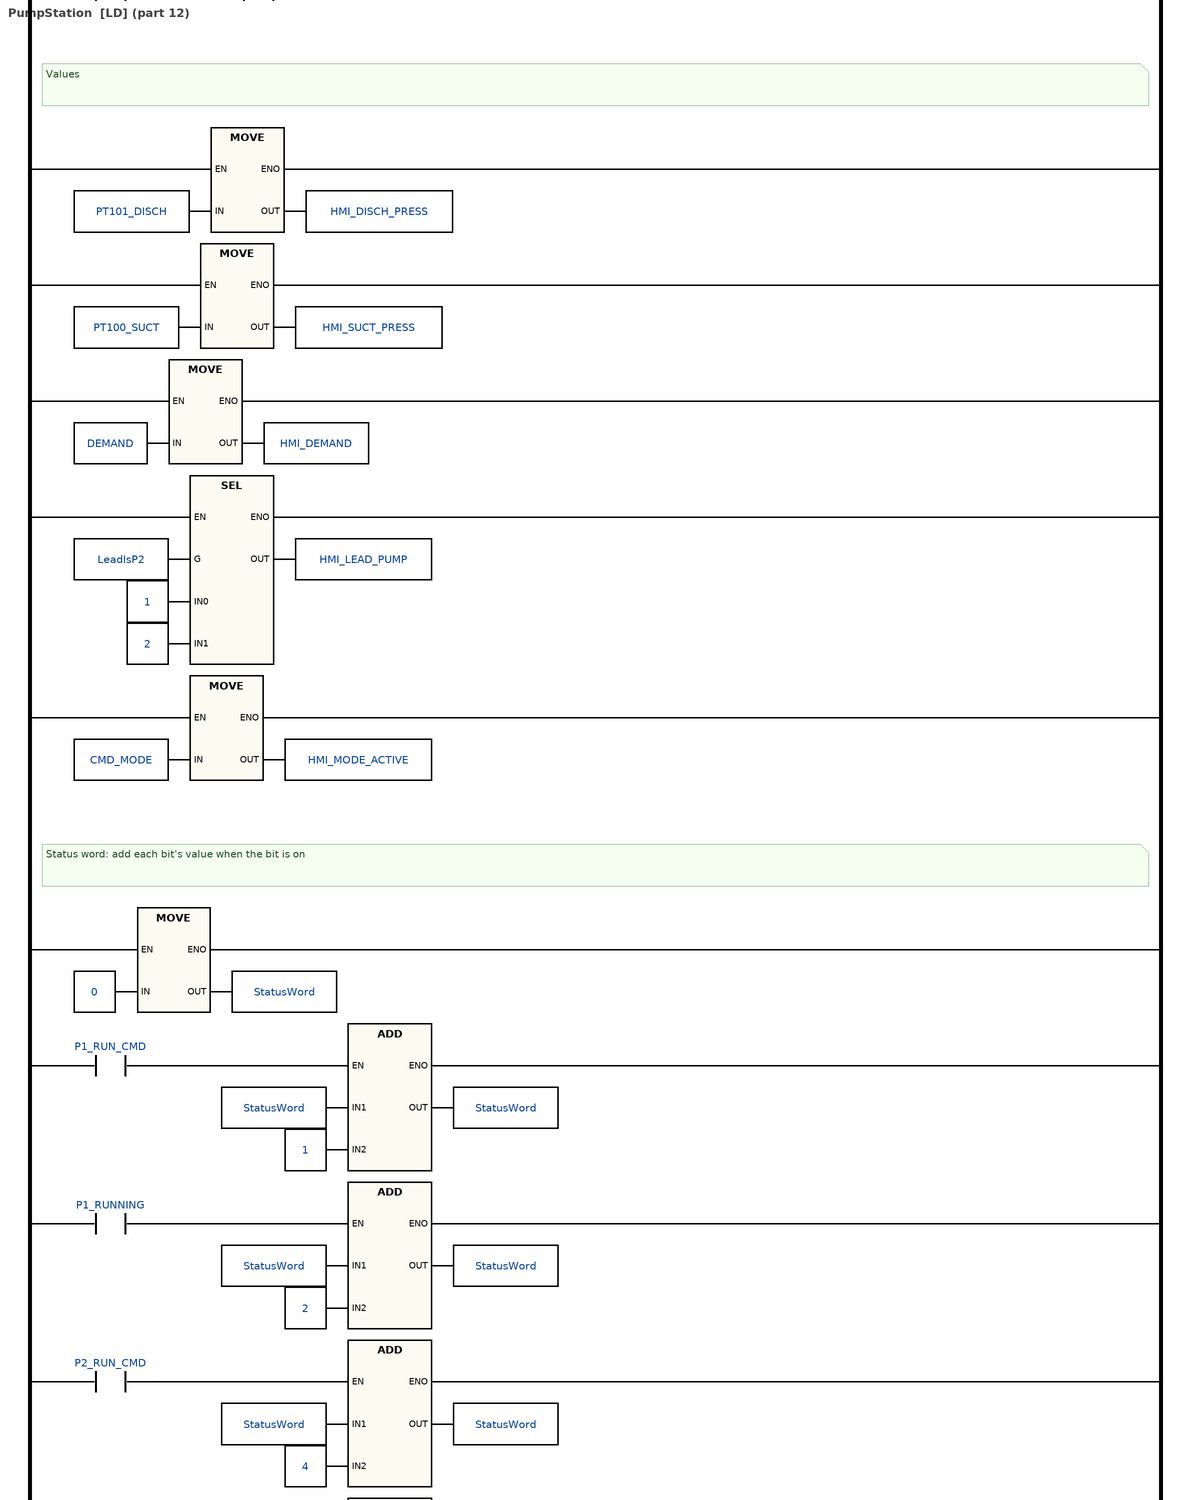
(* Values *)
HMI_DISCH_PRESS := PT101_DISCH;
HMI_SUCT_PRESS := PT100_SUCT;
HMI_DEMAND := DEMAND;
HMI_LEAD_PUMP := SEL(LeadIsP2, 1, 2);
HMI_MODE_ACTIVE := CMD_MODE;
(* Status word: add each bit's value when the bit is on *)
StatusWord := 0;
IF P1_RUN_CMD THEN StatusWord := StatusWord + 1; END_IF;
IF P1_RUNNING THEN StatusWord := StatusWord + 2; END_IF;
IF P2_RUN_CMD THEN StatusWord := StatusWord + 4; END_IF;
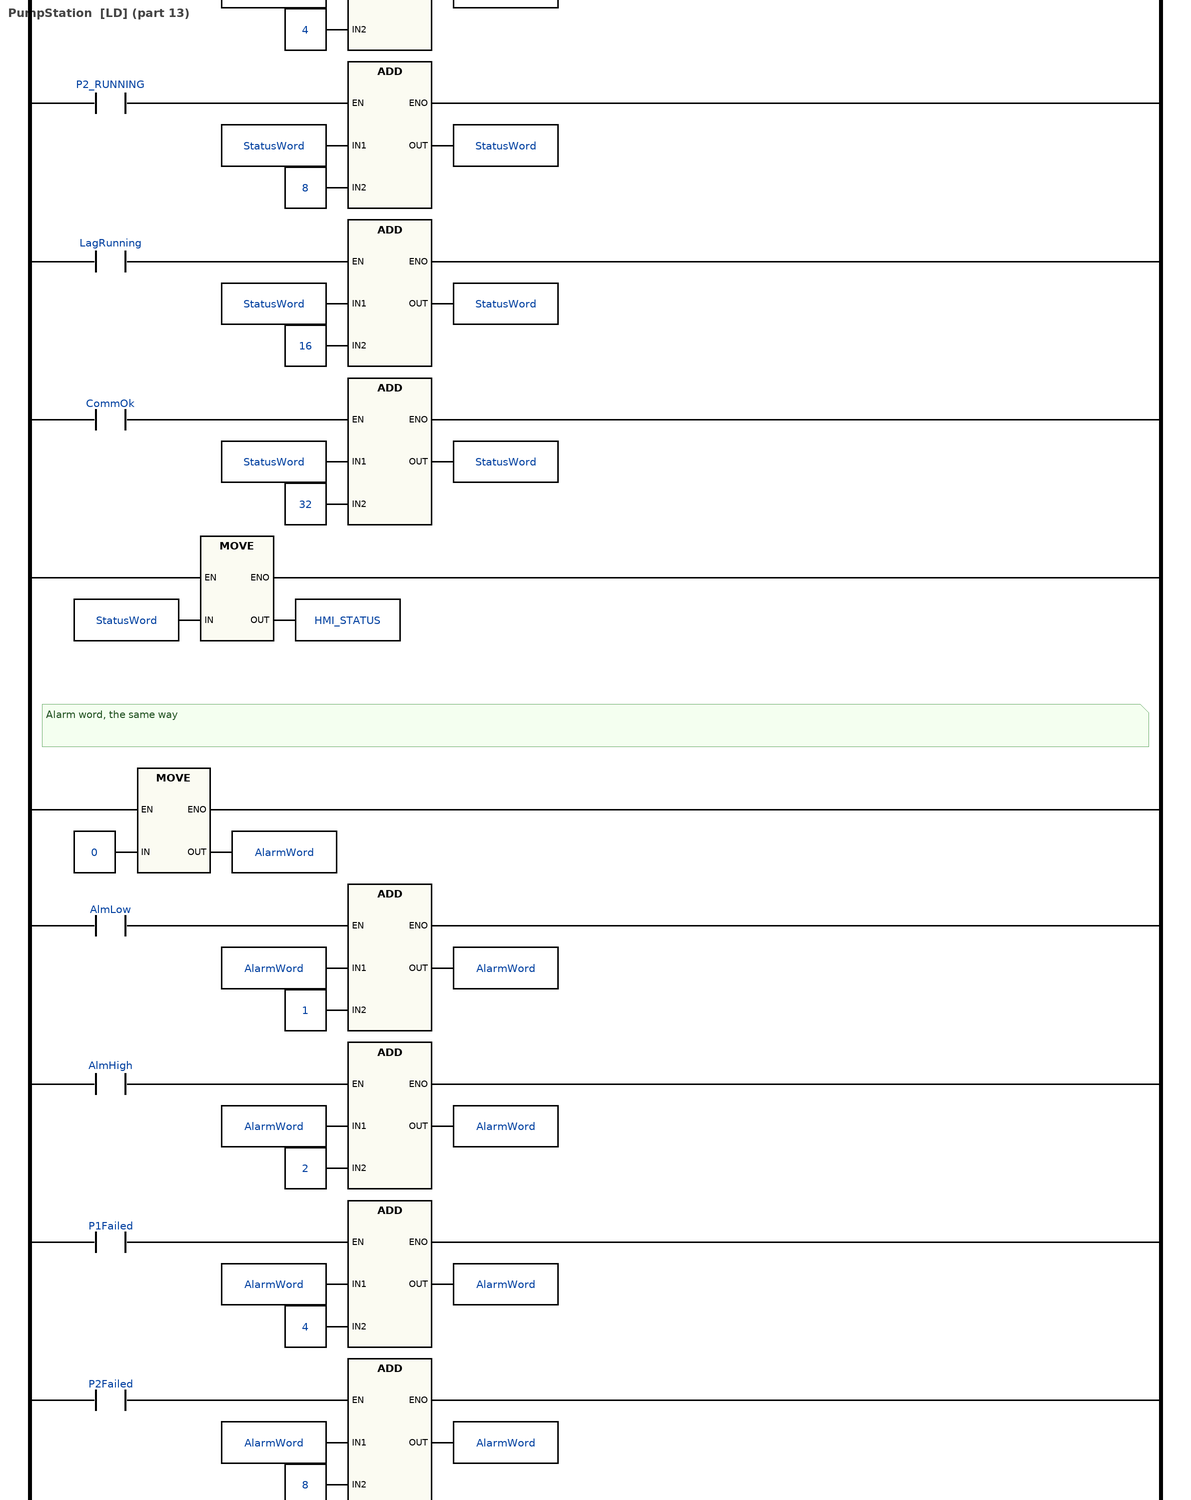
IF P2_RUNNING THEN StatusWord := StatusWord + 8; END_IF;
IF LagRunning THEN StatusWord := StatusWord + 16; END_IF;
IF CommOk THEN StatusWord := StatusWord + 32; END_IF;
HMI_STATUS := StatusWord;
(* Alarm word, the same way *)
AlarmWord := 0;
IF AlmLow THEN AlarmWord := AlarmWord + 1; END_IF;
IF AlmHigh THEN AlarmWord := AlarmWord + 2; END_IF;
IF P1Failed THEN AlarmWord := AlarmWord + 4; END_IF;
IF P2Failed THEN AlarmWord := AlarmWord + 8; END_IF;
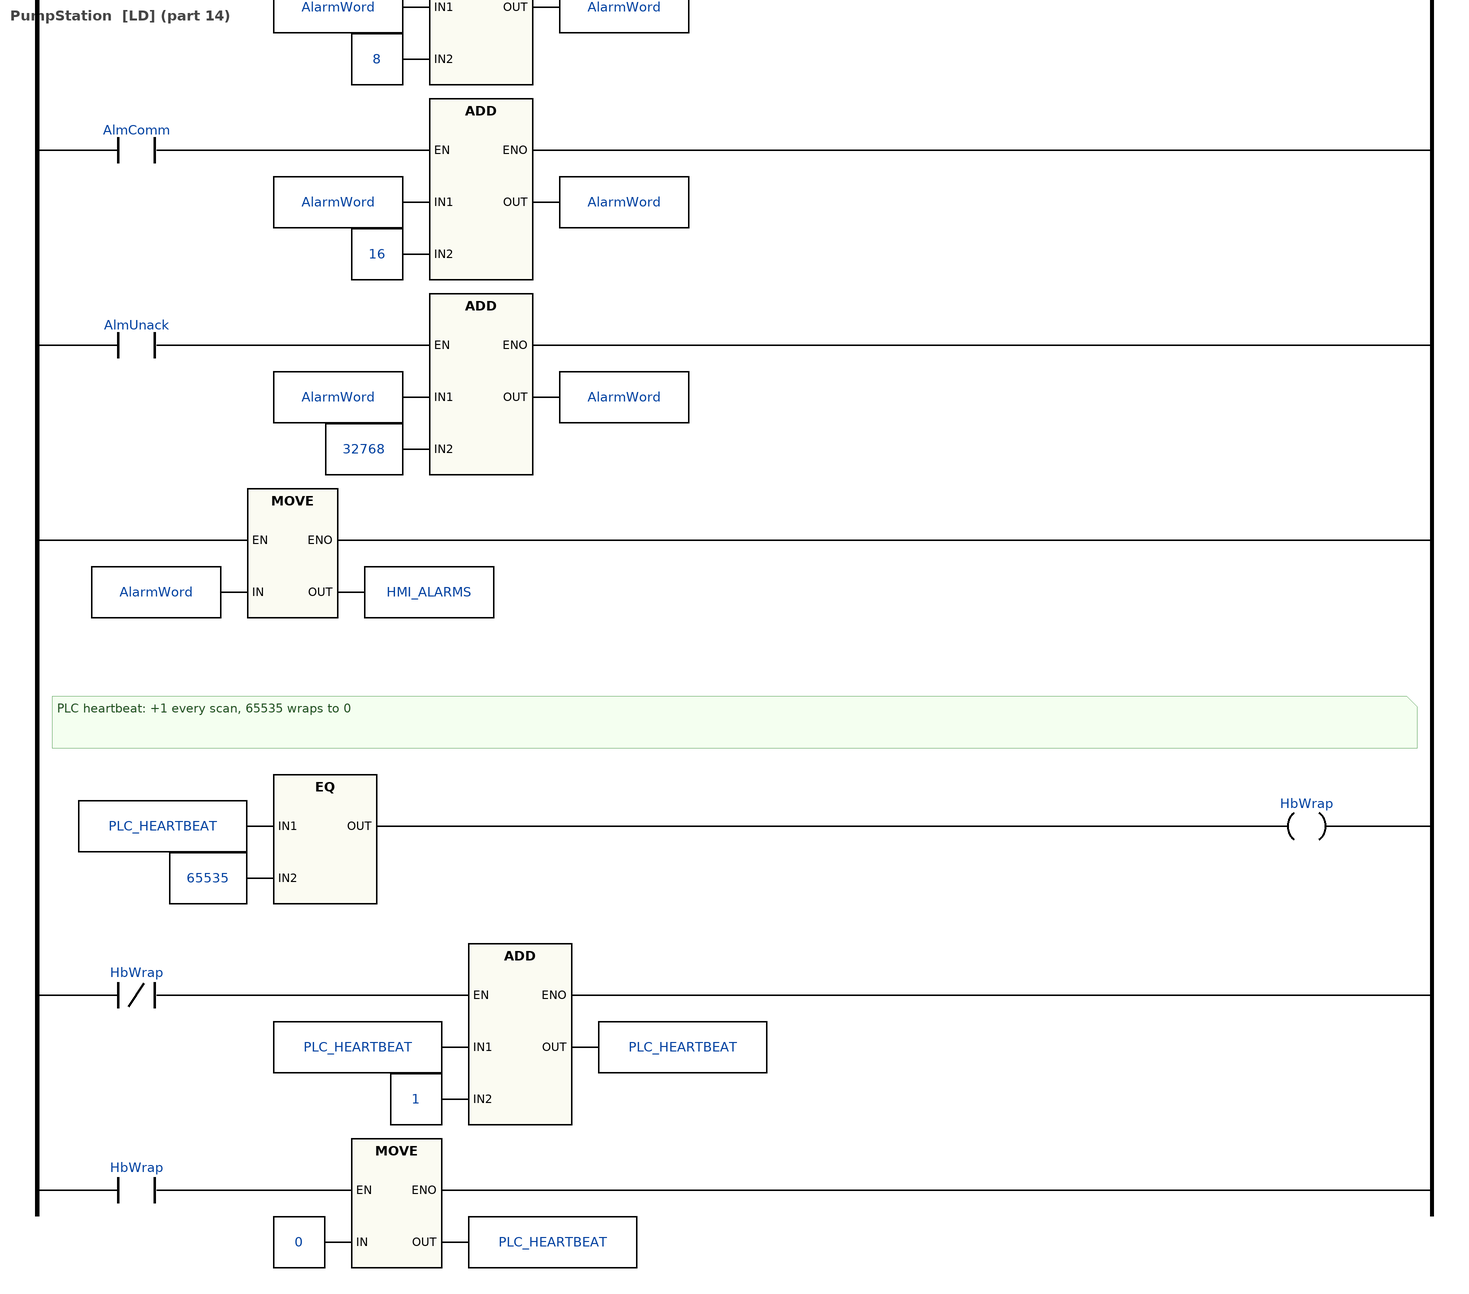
IF AlmComm THEN AlarmWord := AlarmWord + 16; END_IF;
IF AlmUnack THEN AlarmWord := AlarmWord + 32768; END_IF;
HMI_ALARMS := AlarmWord;
(* PLC heartbeat: +1 every scan, 65535 wraps to 0 *)
HbWrap := PLC_HEARTBEAT = 65535;
IF NOT HbWrap THEN PLC_HEARTBEAT := PLC_HEARTBEAT + 1; END_IF;
IF HbWrap THEN PLC_HEARTBEAT := 0; END_IF;
END_PROGRAM

CONFIGURATION Config0
  RESOURCE Res0 ON PLC
    TASK MainTask(INTERVAL := T#100ms, PRIORITY := 0);
    PROGRAM Inst0 WITH MainTask : PumpStation;
  END_RESOURCE
END_CONFIGURATION
